PROGRAM main
  VAR
    MARCHA AT %IX0.0  : BOOL; (* S1, pulsador NA *)
    PARADA AT %IX0.1  : BOOL; (* S2, pulsador NC *)
    TERMICO AT %IX0.2 : BOOL; (* F1, térmico NC *)
    KM1 AT %QX0.0     : BOOL; (* contactor del motor *)
    H1 AT %QX0.1      : BOOL; (* piloto de falla *)
    H2 AT %QX0.2      : BOOL; (* piloto de marcha *)
    FALLA             : BOOL; (* falla del térmico memorizada *)
    RS_KM1            : RS;
    SR_FALLA          : SR;
  END_VAR
  VAR  (* added by the conversion: wires and edge detectors of the diagram *)
    _NOT2_OUT : BOOL;
    _NOT5_OUT : BOOL;
    _AND4_OUT : BOOL;
    _NOT12_OUT : BOOL;
    _AND10_OUT : BOOL;
    _NOT15_OUT : BOOL;
    _NOT17_OUT : BOOL;
    _OR14_OUT : BOOL;
  END_VAR

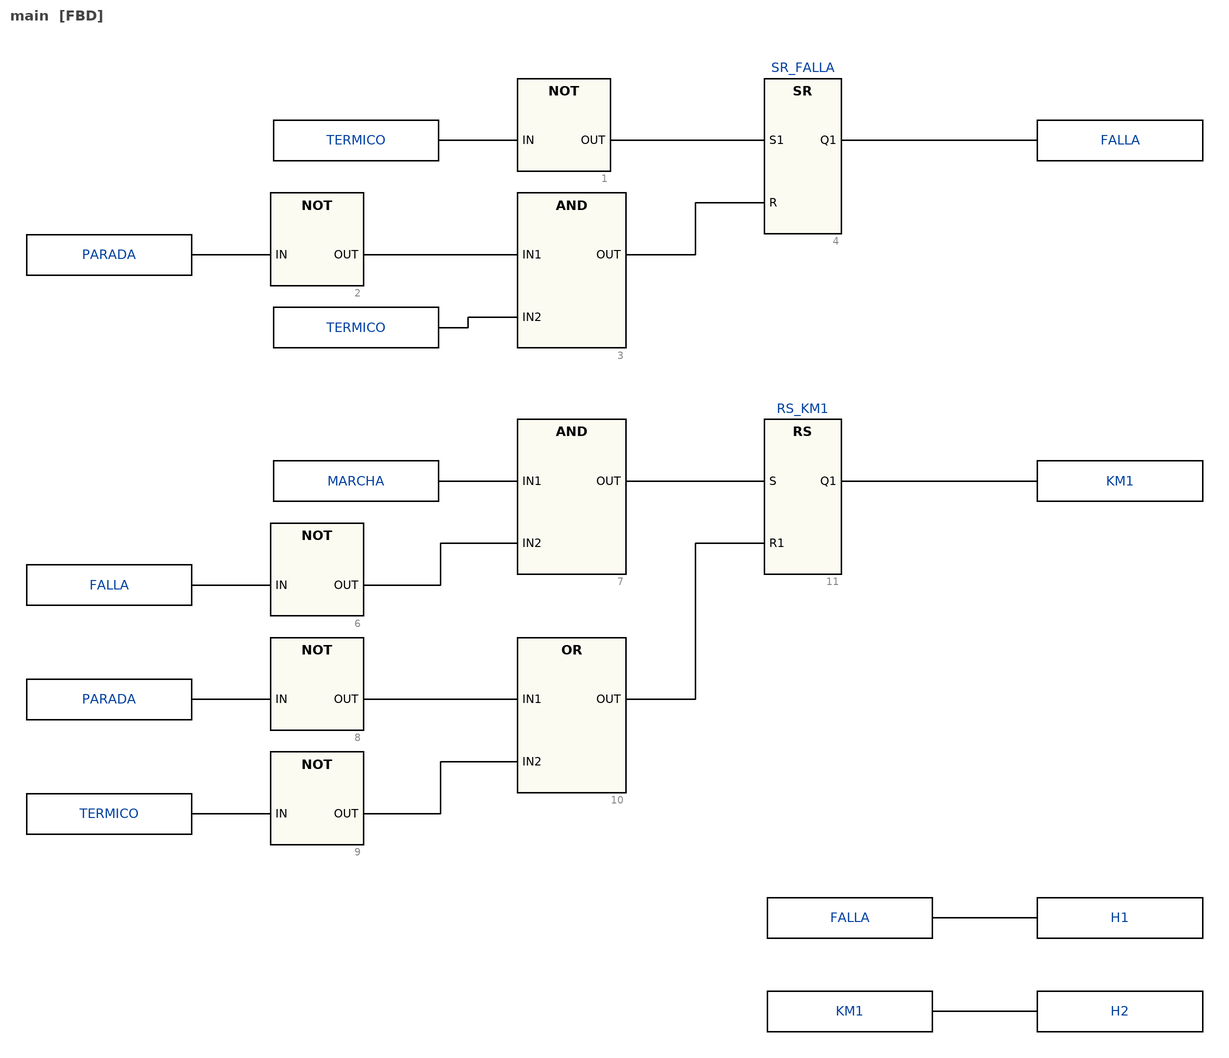
(* FBD diagram, written out as Structured Text *)
_NOT2_OUT := NOT TERMICO;
_NOT5_OUT := NOT PARADA;
_AND4_OUT := _NOT5_OUT AND TERMICO;
SR_FALLA(S1 := _NOT2_OUT, R := _AND4_OUT);
FALLA := SR_FALLA.Q1;
_NOT12_OUT := NOT FALLA;
_AND10_OUT := MARCHA AND _NOT12_OUT;
_NOT15_OUT := NOT PARADA;
_NOT17_OUT := NOT TERMICO;
_OR14_OUT := _NOT15_OUT OR _NOT17_OUT;
RS_KM1(S := _AND10_OUT, R1 := _OR14_OUT);
KM1 := RS_KM1.Q1;
H1 := FALLA;
H2 := KM1;
END_PROGRAM
